(* IEC 61131-3 sources: plc-vscode/tests/st/test-ready/trust-platform/examples/OSCAT/kiln_dryer_decorator_strategy/oop/src, 3 files *)

(* ---- Main.st ---- *)
(* Pattern role: IMoistureSource is the contract boundary for the Decorator and Strategy example. *)
INTERFACE IMoistureSource
    PROPERTY Value : REAL
    GET
    END_GET
    END_PROPERTY
    PROPERTY Quality : BYTE
    GET
    END_GET
    END_PROPERTY
    METHOD Update
    END_METHOD
END_INTERFACE

(* Pattern role: IDryingStrategy is the contract boundary for the Decorator and Strategy example. *)
INTERFACE IDryingStrategy
    PROPERTY ProfileId : INT
    GET
    END_GET
    END_PROPERTY
    METHOD HeatCommand : REAL
    VAR_INPUT
        MoisturePct : REAL;
    END_VAR
    END_METHOD
    METHOD FanSpeed : REAL
    VAR_INPUT
        MoisturePct : REAL;
    END_VAR
    END_METHOD
END_INTERFACE

(* Pattern role: RawMoistureInput is a concrete implementation in the Decorator and Strategy example. *)
FUNCTION_BLOCK RawMoistureInput IMPLEMENTS IMoistureSource
VAR
    ValueValue : REAL;
    QualityValue : BYTE := BYTE#2;
END_VAR
METHOD PUBLIC SetRaw
VAR_INPUT
    MoisturePct : REAL;
END_VAR
ValueValue := MoisturePct;
END_METHOD
METHOD PUBLIC Update
END_METHOD
PUBLIC PROPERTY Value : REAL
GET
    Value := ValueValue;
END_GET
END_PROPERTY
PUBLIC PROPERTY Quality : BYTE
GET
    Quality := QualityValue;
END_GET
END_PROPERTY
END_FUNCTION_BLOCK

(* Pattern role: MoistureClampDecorator is a concrete implementation in the Decorator and Strategy example. *)
FUNCTION_BLOCK MoistureClampDecorator IMPLEMENTS IMoistureSource
VAR
    Inner : IMoistureSource;
    ValueValue : REAL;
    QualityValue : BYTE;
END_VAR
METHOD PUBLIC Wrap
VAR_INPUT
    Source : IMoistureSource;
END_VAR
Inner := Source;
END_METHOD
METHOD PUBLIC Update
Inner.Update();
IF Inner.Value < REAL#0.0 THEN
    ValueValue := REAL#0.0;
    QualityValue := BYTE#0;
ELSIF Inner.Value > REAL#100.0 THEN
    ValueValue := REAL#100.0;
    QualityValue := BYTE#0;
ELSE
    ValueValue := Inner.Value;
    QualityValue := Inner.Quality;
END_IF;
END_METHOD
PUBLIC PROPERTY Value : REAL
GET
    Value := ValueValue;
END_GET
END_PROPERTY
PUBLIC PROPERTY Quality : BYTE
GET
    Quality := QualityValue;
END_GET
END_PROPERTY
END_FUNCTION_BLOCK

(* Pattern role: MoistureFilterDecorator is a concrete implementation in the Decorator and Strategy example. *)
FUNCTION_BLOCK MoistureFilterDecorator IMPLEMENTS IMoistureSource
VAR
    Inner : IMoistureSource;
    Filter : Pt1Filter;
    ValueValue : REAL;
    QualityValue : BYTE;
END_VAR
METHOD PUBLIC Wrap
VAR_INPUT
    Source : IMoistureSource;
END_VAR
Inner := Source;
Filter.Initialize();
Filter.Configure(TimeConstant := T#1s, Gain := REAL#1.0);
END_METHOD
METHOD PUBLIC Update
Inner.Update();
IF Inner.Quality = BYTE#2 THEN
    ValueValue := Filter.Update(Sample := Inner.Value);
ELSE
    ValueValue := Inner.Value;
END_IF;
QualityValue := Inner.Quality;
END_METHOD
PUBLIC PROPERTY Value : REAL
GET
    Value := ValueValue;
END_GET
END_PROPERTY
PUBLIC PROPERTY Quality : BYTE
GET
    Quality := QualityValue;
END_GET
END_PROPERTY
END_FUNCTION_BLOCK

(* Pattern role: SoftwoodStrategy is a concrete implementation in the Decorator and Strategy example. *)
FUNCTION_BLOCK SoftwoodStrategy IMPLEMENTS IDryingStrategy
METHOD PUBLIC HeatCommand : REAL
VAR_INPUT
    MoisturePct : REAL;
END_VAR
HeatCommand := LIMIT(REAL#0.0, (MoisturePct - REAL#12.0) * REAL#3.0, REAL#100.0);
END_METHOD
METHOD PUBLIC FanSpeed : REAL
VAR_INPUT
    MoisturePct : REAL;
END_VAR
FanSpeed := REAL#45.0;
END_METHOD
PUBLIC PROPERTY ProfileId : INT
GET
    ProfileId := INT#1;
END_GET
END_PROPERTY
END_FUNCTION_BLOCK

(* Pattern role: HardwoodStrategy is a concrete implementation in the Decorator and Strategy example. *)
FUNCTION_BLOCK HardwoodStrategy IMPLEMENTS IDryingStrategy
METHOD PUBLIC HeatCommand : REAL
VAR_INPUT
    MoisturePct : REAL;
END_VAR
HeatCommand := LIMIT(REAL#0.0, (MoisturePct - REAL#8.0) * REAL#2.0, REAL#80.0);
END_METHOD
METHOD PUBLIC FanSpeed : REAL
VAR_INPUT
    MoisturePct : REAL;
END_VAR
FanSpeed := REAL#30.0;
END_METHOD
PUBLIC PROPERTY ProfileId : INT
GET
    ProfileId := INT#2;
END_GET
END_PROPERTY
END_FUNCTION_BLOCK

(* Composition role: KilnDryerController owns the collaborating objects used by this Decorator and Strategy example. *)
FUNCTION_BLOCK KilnDryerController
VAR
    Raw : RawMoistureInput;
    Clamped : MoistureClampDecorator;
    Filtered : MoistureFilterDecorator;
    Moisture : IMoistureSource;
    Softwood : SoftwoodStrategy;
    Hardwood : HardwoodStrategy;
    ActiveStrategy : IDryingStrategy;
    ActiveProfileIdValue : INT;
    HeatCommandValue : REAL;
    FanSpeedValue : REAL;
END_VAR
METHOD PUBLIC Initialize
Clamped.Wrap(Source := Raw);
Filtered.Wrap(Source := Clamped);
Moisture := Filtered;
ActiveStrategy := Softwood;
END_METHOD
METHOD PUBLIC Update : REAL
VAR_INPUT
    ProductId : INT;
    RawMoisturePct : REAL;
END_VAR
Raw.SetRaw(MoisturePct := RawMoisturePct);
IF ProductId = INT#2 THEN ActiveStrategy := Hardwood; ELSE ActiveStrategy := Softwood; END_IF;
Moisture.Update();
ActiveProfileIdValue := ActiveStrategy.ProfileId;
HeatCommandValue := ActiveStrategy.HeatCommand(MoisturePct := Moisture.Value);
FanSpeedValue := ActiveStrategy.FanSpeed(MoisturePct := Moisture.Value);
Update := HeatCommandValue;
END_METHOD
PUBLIC PROPERTY ActiveProfileId : INT
GET
    ActiveProfileId := ActiveProfileIdValue;
END_GET
END_PROPERTY
PUBLIC PROPERTY HeatCommand : REAL
GET
    HeatCommand := HeatCommandValue;
END_GET
END_PROPERTY
PUBLIC PROPERTY FanSpeed : REAL
GET
    FanSpeed := FanSpeedValue;
END_GET
END_PROPERTY
PUBLIC PROPERTY ConditionedMoisture : REAL
GET
    ConditionedMoisture := Moisture.Value;
END_GET
END_PROPERTY
PUBLIC PROPERTY MoistureQuality : BYTE
GET
    MoistureQuality := Moisture.Quality;
END_GET
END_PROPERTY
END_FUNCTION_BLOCK

(* Scan role: Main wires the example objects and exposes the PLC call path under test. *)
PROGRAM Main
VAR
    Dryer : KilnDryerController;
    ProductId : INT;
    MoistureRaw : INT;
    HeatCommandRaw : INT;
    FanSpeedRaw : INT;
END_VAR
Dryer.Initialize();
HeatCommandRaw := REAL_TO_INT(Dryer.Update(ProductId := ProductId, RawMoisturePct := INT_TO_REAL(MoistureRaw) / REAL#10.0));
FanSpeedRaw := REAL_TO_INT(Dryer.FanSpeed);
END_PROGRAM

(* ---- Configuration.st ---- *)
CONFIGURATION KilnDryerDecoratorStrategyOopConfiguration
RESOURCE Cpu0 ON PLC
    TASK MainTask (INTERVAL := T#100ms, PRIORITY := 1);
    PROGRAM Dryer WITH MainTask : Main;
END_RESOURCE
VAR_CONFIG
    Dryer.ProductId AT %IW0 : INT;
    Dryer.MoistureRaw AT %IW2 : INT;
    Dryer.HeatCommandRaw AT %QW0 : INT;
    Dryer.FanSpeedRaw AT %QW2 : INT;
END_VAR
END_CONFIGURATION

(* ---- Tests.st ---- *)
TEST_PROGRAM KilnDecoratorClampsBadMoisture
VAR
    Dryer : KilnDryerController;
    Heat : REAL;
END_VAR
Dryer.Initialize();
Heat := Dryer.Update(ProductId := INT#1, RawMoisturePct := REAL#120.0);
ASSERT_EQUAL(EXPECTED := BYTE#0, ACTUAL := Dryer.MoistureQuality);
ASSERT_NEAR(EXPECTED := REAL#100.0, ACTUAL := Dryer.ConditionedMoisture, DELTA := REAL#0.001);
END_TEST_PROGRAM

TEST_PROGRAM KilnStrategiesSelectDifferentFanSpeed
VAR
    Dryer : KilnDryerController;
    SoftFan : REAL;
    HardFan : REAL;
END_VAR
Dryer.Initialize();
Dryer.Update(ProductId := INT#1, RawMoisturePct := REAL#20.0);
SoftFan := Dryer.FanSpeed;
Dryer.Update(ProductId := INT#2, RawMoisturePct := REAL#20.0);
HardFan := Dryer.FanSpeed;
ASSERT_TRUE(IN := SoftFan > HardFan);
ASSERT_EQUAL(EXPECTED := INT#2, ACTUAL := Dryer.ActiveProfileId);
END_TEST_PROGRAM

(* Decorator + strategy combined-flow test: drives a sequence of bad
   inputs (clamped) -> good inputs (passes through) -> profile switch
   on the same instance. Catches bugs where the decorator's quality
   flag stays bad after a clean reading, or where strategy selection
   doesn't re-evaluate when ProductId changes. *)
TEST_PROGRAM KilnDecoratorAndStrategyReevaluateAcrossScans
VAR
    Dryer : KilnDryerController;
END_VAR

Dryer.Initialize();

(* Bad input - quality clamped *)
Dryer.Update(ProductId := INT#1, RawMoisturePct := REAL#120.0);
ASSERT_EQUAL(EXPECTED := BYTE#0, ACTUAL := Dryer.MoistureQuality);

(* Recover - quality must report good *)
Dryer.Update(ProductId := INT#1, RawMoisturePct := REAL#22.0);
ASSERT_EQUAL(EXPECTED := BYTE#2, ACTUAL := Dryer.MoistureQuality);

(* Switch product (Strategy change) on recovered signal *)
Dryer.Update(ProductId := INT#2, RawMoisturePct := REAL#22.0);
ASSERT_EQUAL(EXPECTED := INT#2, ACTUAL := Dryer.ActiveProfileId);

(* Switch back to product 1 - profile must follow *)
Dryer.Update(ProductId := INT#1, RawMoisturePct := REAL#22.0);
ASSERT_EQUAL(EXPECTED := INT#1, ACTUAL := Dryer.ActiveProfileId);
END_TEST_PROGRAM

(* Boundary test: clamp must trip on the negative side too. A negative
   moisture reading is physically impossible and must not be passed
   through. *)
TEST_PROGRAM KilnDecoratorClampsNegativeMoisture
VAR
    Dryer : KilnDryerController;
END_VAR
Dryer.Initialize();
Dryer.Update(ProductId := INT#1, RawMoisturePct := REAL#-5.0);
ASSERT_EQUAL(EXPECTED := BYTE#0, ACTUAL := Dryer.MoistureQuality);
ASSERT_NEAR(EXPECTED := REAL#0.0, ACTUAL := Dryer.ConditionedMoisture, DELTA := REAL#0.001);
(* Heat command must be zero because (clamped 0 - 12 setpoint) * gain
   limits to zero on the lower bound *)
ASSERT_NEAR(EXPECTED := REAL#0.0, ACTUAL := Dryer.HeatCommand, DELTA := REAL#0.001);
END_TEST_PROGRAM

(* Strategy edge inputs: each strategy maps the moisture-vs-target
   curve to a heat command. Below target, heat is zero; above target,
   it grows linearly until the per-strategy ceiling. *)
TEST_PROGRAM KilnStrategiesRespectTargetAndCeilings
VAR
    Soft : SoftwoodStrategy;
    Hard : HardwoodStrategy;
END_VAR

(* Softwood target 12, gain 3, ceiling 100 *)
ASSERT_NEAR(EXPECTED := REAL#0.0, ACTUAL := Soft.HeatCommand(MoisturePct := REAL#10.0), DELTA := REAL#0.001);
ASSERT_NEAR(EXPECTED := REAL#0.0, ACTUAL := Soft.HeatCommand(MoisturePct := REAL#12.0), DELTA := REAL#0.001);
ASSERT_NEAR(EXPECTED := REAL#15.0, ACTUAL := Soft.HeatCommand(MoisturePct := REAL#17.0), DELTA := REAL#0.001);
(* Saturation: above 12 + 100/3 = 45.33 the ceiling clips *)
ASSERT_NEAR(EXPECTED := REAL#100.0, ACTUAL := Soft.HeatCommand(MoisturePct := REAL#80.0), DELTA := REAL#0.001);

(* Hardwood target 8, gain 2, ceiling 80 *)
ASSERT_NEAR(EXPECTED := REAL#0.0, ACTUAL := Hard.HeatCommand(MoisturePct := REAL#5.0), DELTA := REAL#0.001);
ASSERT_NEAR(EXPECTED := REAL#0.0, ACTUAL := Hard.HeatCommand(MoisturePct := REAL#8.0), DELTA := REAL#0.001);
ASSERT_NEAR(EXPECTED := REAL#10.0, ACTUAL := Hard.HeatCommand(MoisturePct := REAL#13.0), DELTA := REAL#0.001);
(* Hardwood ceiling: above 8 + 80/2 = 48 the ceiling clips *)
ASSERT_NEAR(EXPECTED := REAL#80.0, ACTUAL := Hard.HeatCommand(MoisturePct := REAL#60.0), DELTA := REAL#0.001);

(* Per-product fan speed *)
ASSERT_NEAR(EXPECTED := REAL#45.0, ACTUAL := Soft.FanSpeed(MoisturePct := REAL#20.0), DELTA := REAL#0.001);
ASSERT_NEAR(EXPECTED := REAL#30.0, ACTUAL := Hard.FanSpeed(MoisturePct := REAL#20.0), DELTA := REAL#0.001);
END_TEST_PROGRAM

(* Decorator chain isolation: two RawMoistureInput sources can each
   feed an independent clamp without bleeding. The pattern requires
   one wrap per source; two wraps must be independent. *)
TEST_PROGRAM KilnDecoratorChainsAreIndependent
VAR
    SourceA : RawMoistureInput;
    SourceB : RawMoistureInput;
    ClampA : MoistureClampDecorator;
    ClampB : MoistureClampDecorator;
END_VAR

ClampA.Wrap(Source := SourceA);
ClampB.Wrap(Source := SourceB);

SourceA.SetRaw(MoisturePct := REAL#150.0);
SourceB.SetRaw(MoisturePct := REAL#22.0);
ClampA.Update();
ClampB.Update();

(* A is clamped, B is in range *)
ASSERT_NEAR(EXPECTED := REAL#100.0, ACTUAL := ClampA.Value, DELTA := REAL#0.001);
ASSERT_EQUAL(EXPECTED := BYTE#0, ACTUAL := ClampA.Quality);
ASSERT_NEAR(EXPECTED := REAL#22.0, ACTUAL := ClampB.Value, DELTA := REAL#0.001);
ASSERT_EQUAL(EXPECTED := BYTE#2, ACTUAL := ClampB.Quality);

(* Drive A back into range and B out: the flags must follow each
   independently *)
SourceA.SetRaw(MoisturePct := REAL#30.0);
SourceB.SetRaw(MoisturePct := REAL#-10.0);
ClampA.Update();
ClampB.Update();
ASSERT_EQUAL(EXPECTED := BYTE#2, ACTUAL := ClampA.Quality);
ASSERT_EQUAL(EXPECTED := BYTE#0, ACTUAL := ClampB.Quality);
ASSERT_NEAR(EXPECTED := REAL#0.0, ACTUAL := ClampB.Value, DELTA := REAL#0.001);
END_TEST_PROGRAM
